FUNCTION_BLOCK FB_Samples
VAR_INPUT
    index : INT := 1;
    value : REAL;
    write : BOOL;
END_VAR
VAR_OUTPUT
    values : ARRAY[1..3] OF REAL := [3(0.0)];
END_VAR

IF write THEN
    values[index] := value;
END_IF;

END_FUNCTION_BLOCK

(* stored: Version 1.1.0.1 *)
